// TIA Portal V19 export
VAR_GLOBAL   // PLC tag table "Power"
   DI_MainSupply_Ok AT %I0.2 : Bool;
   DI_PowerSupply_OK AT %I0.3 : Bool;
END_VAR
